PROGRAM main
  VAR
    oscillator AT %IX0.0 : BOOL;
    full_up AT %QX0.0 : BOOL;
    full_down AT %QX0.1 : BOOL;
    ramp_cnt : INT;
    CTUD0 : CTUD;
  END_VAR

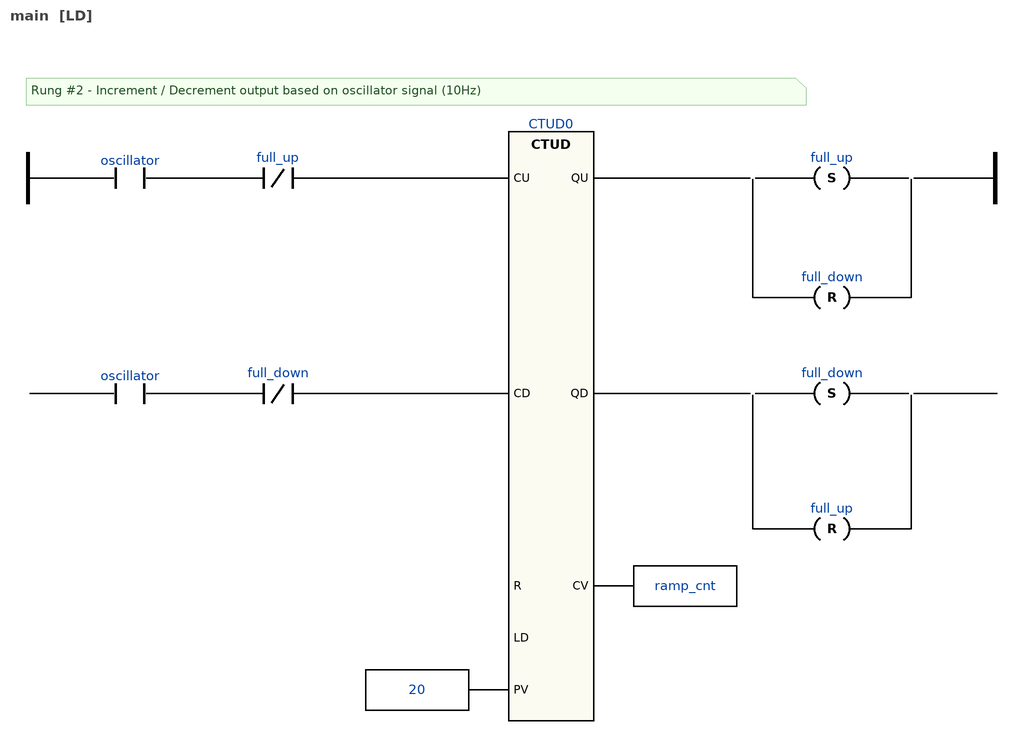
(* LD diagram, written out as Structured Text *)
(* Rung #2 - Increment / Decrement output based on oscillator signal (10Hz) *)
CTUD0(CU := oscillator AND NOT full_up, CD := oscillator AND NOT full_down, PV := 20);
IF CTUD0.QU THEN full_up := TRUE; END_IF;
IF CTUD0.QU THEN full_down := FALSE; END_IF;
IF CTUD0.QD THEN full_down := TRUE; END_IF;
IF CTUD0.QD THEN full_up := FALSE; END_IF;
ramp_cnt := CTUD0.CV;
END_PROGRAM
